// TIA Portal V20 export
TYPE "WT2_Vd_Status_2_UDT"
   STRUCT
      iHandshake : Int;
      Fehler : Struct
         bE0128_Reserviert : Bool;
         bE0129_Reserviert : Bool;
         bE0130_Reserviert : Bool;
         bE0131_Reserviert : Bool;
         bE0132_Reserviert : Bool;
         bE0133_Reserviert : Bool;
         bE0134_Reserviert : Bool;
         bE0135_Reserviert : Bool;
         bE0136_Reserviert : Bool;
         bE0137_Reserviert : Bool;
         bE0138_VorschmNoetig : Bool;
         bE0139_KonfigFehlerHaltebetr : Bool;
         bE0140_FehlerTTOPHKZuTief : Bool;
         bE0141_FehlerTTOPHKZuHoch : Bool;
         bE0142_KonfigFehlerKeinDefVi : Bool;
         b37_Reserve : Bool;
         by04_Reserve : Byte;
         by05_Reserve : Byte;
         by06_Reserve : Byte;
         by07_Reserve : Byte;
         by08_Reserve : Byte;
         by09_Reserve : Byte;
         by10_Reserve : Byte;
         by11_Reserve : Byte;
         by12_Reserve : Byte;
         by13_Reserve : Byte;
         by14_Reserve : Byte;
         by15_Reserve : Byte;
         by16_Reserve : Byte;
         by17_Reserve : Byte;
      END_STRUCT;
      Alarm : Struct
         bA1128_Vorschm3Tagen : Bool;
         bA1129_Vorschm2Tagen : Bool;
         bA1130_Vorschm1Tag : Bool;
         bA1131_Reserviert : Bool;
         bA1132_Reserviert : Bool;
         bA1133_Reserviert : Bool;
         bA1134_Reserviert : Bool;
         bA1135_Reserviert : Bool;
         bA1136_Reserviert : Bool;
         bA1137_Reserviert : Bool;
         bA1138_Reserviert : Bool;
         bA1139_Reserviert : Bool;
         bA1140_AlarmTTOPHKZuTief : Bool;
         bA1141_AlarmTTOPHKZuHoch : Bool;
         bA1142_Reserviert : Bool;
         b197_Reserve : Bool;
         by20_Reserve : Byte;
         by21_Reserve : Byte;
         by22_Reserve : Byte;
         by23_Reserve : Byte;
         by24_Reserve : Byte;
         by25_Reserve : Byte;
         by26_Reserve : Byte;
         by27_Reserve : Byte;
         by28_Reserve : Byte;
         by29_Reserve : Byte;
         by30_Reserve : Byte;
         by31_Reserve : Byte;
         by32_Reserve : Byte;
         by33_Reserve : Byte;
      END_STRUCT;
      Zustand : Struct
         by34_Reserve : Byte;
         by35_Reserve : Byte;
         by36_Reserve : Byte;
         by37_Reserve : Byte;
         by38_Reserve : Byte;
         by39_Reserve : Byte;
         by40_Reserve : Byte;
         by41_Reserve : Byte;
         by42_Reserve : Byte;
         by43_Reserve : Byte;
         by44_Reserve : Byte;
         by45_Reserve : Byte;
      END_STRUCT;
      DigIn : Struct
         by46_Reserve : Byte;
         by47_Reserve : Byte;
         by48_Reserve : Byte;
         by49_Reserve : Byte;
         by50_Reserve : Byte;
         by51_Reserve : Byte;
         by52_Reserve : Byte;
         by53_Reserve : Byte;
      END_STRUCT;
      DigOut : Struct
         by54_Reserve : Byte;
         by55_Reserve : Byte;
         by56_Reserve : Byte;
         by57_Reserve : Byte;
         by58_Reserve : Byte;
         by59_Reserve : Byte;
         by60_Reserve : Byte;
         by61_Reserve : Byte;
      END_STRUCT;
      rNDAbscheiderNiveau : Real;
      rEconomiserNiveau : Real;
      rTVerdichterkühlAustritt : Real;
      rTZwStufeSaugHD : Real;
      rTEconomiser : Real;
      rTTOPHeizenKühlen : Real;
      rEconomiserAnalog : Real;
      rUeberhitzungsventil : Real;
      rAnlaufentlastungAnalog : Real;
      rOelpumpenAusgang : Real;
      rEcoNiveaureglerAusgang : Real;
      diLaeuftSeit : DInt;
      rCPos : Real;
      rReserveReal : Array[0..215] of Real;
   END_STRUCT;
END_TYPE
